TYPE "ST_ShiftCalendarV3"
VERSION : 0.1
   STRUCT
      "SchemaVersion" : UInt;
      "UtcOffsetMin" : DInt;
      "Rows" : Array[1..5] of "ST_ShiftRowV3";
   END_STRUCT;
END_TYPE
